// TIA Portal V21 export
// export: Created 2026-10-23T20:44:38.1986875Z, ExportSetting WithDefaults, DisplayName Totally Integrated Automation Portal, DisplayVersion V21 Update 1, DisplayName SINAMICS Startdrive Advanced, DisplayVersion V21 HF2, DisplayName SINAMICS Startdrive G110M, G120, G120C, G120D, G120P, G115D, DisplayVersion V21 HF2, DisplayName SINAMICS Startdrive G130, G150, S120, S150, G200, G220, S200, S210, S220, Innomotics MVD, DisplayVersion V21 HF2, DisplayName STEP 7 Professional, DisplayVersion V21 Update 1, DisplayName STEP 7 Safety, DisplayVersion V21, DisplayName Tech WebApplication, DisplayVersion V21, DisplayName WinCC Basic/Comfort/Advanced, DisplayVersion V21 Update 1, DisplayName WinCC Unified, DisplayVersion V21 Update 1
FUNCTION_BLOCK "FB_Doser"   // FB6, SCL
VERSION : 0.1
// stored: Access Published, AutoNumber true, IsIECCheckEnabled false, IsRetainMemResEnabled false, MemoryReserve 100, Namespace Dosing, SetENOAutomatically false, UDAEnableTagReadback false
   VAR_INPUT
      Start : Bool;   // Start dosing
      Stop : Bool;   // Stop dosing
   END_VAR
   VAR_OUTPUT
      Dosing : Bool;   // Dosing is running
      Done : Bool;   // Dosing finished
   END_VAR
   VAR
      Filler { S7_SetPoint := 'True'} : "Filling.FB_Filler";   // Filler of the unit Filling
      Recipe { S7_SetPoint := 'True'} : "Filling.UDT_FillRecipe";   // Recipe of the unit Filling
   END_VAR
BEGIN

       REGION Dosing through the filler
           #Recipe.TargetVolume := 0.5;
           #Filler(Start := #Start, Stop := #Stop, Recipe := #Recipe);
           #Dosing := #Filler.Filling;
           #Done := #Filler.Done;
       END_REGION
END_FUNCTION_BLOCK
